PROGRAM main
  VAR
    SA1 AT %IX0.0 : BOOL; (* mano izquierda *)
    SA2 AT %IX0.1 : BOOL; (* mano derecha *)
    SA3 AT %IX0.2 : BOOL; (* tercera mano *)
    H1 AT %QX0.0  : BOOL; (* prensa *)
    H2 AT %QX0.1  : BOOL;
    H3 AT %QX0.2  : BOOL;
    H5 AT %QX0.4  : BOOL;
  END_VAR

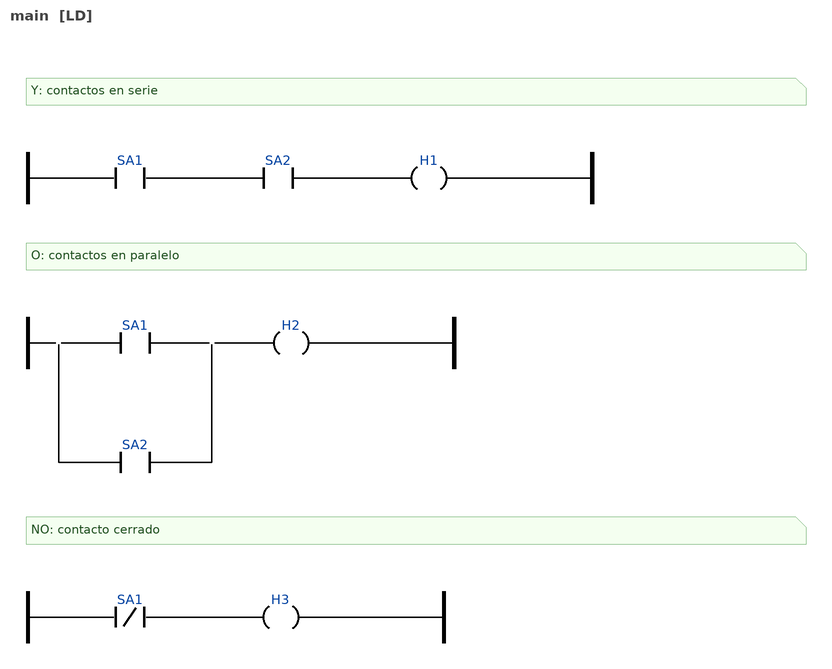
(* LD diagram, written out as Structured Text *)
(* Y: contactos en serie *)
H1 := SA1 AND SA2;
(* O: contactos en paralelo *)
H2 := SA1 OR SA2;
(* NO: contacto cerrado *)
H3 := NOT SA1;
END_PROGRAM
